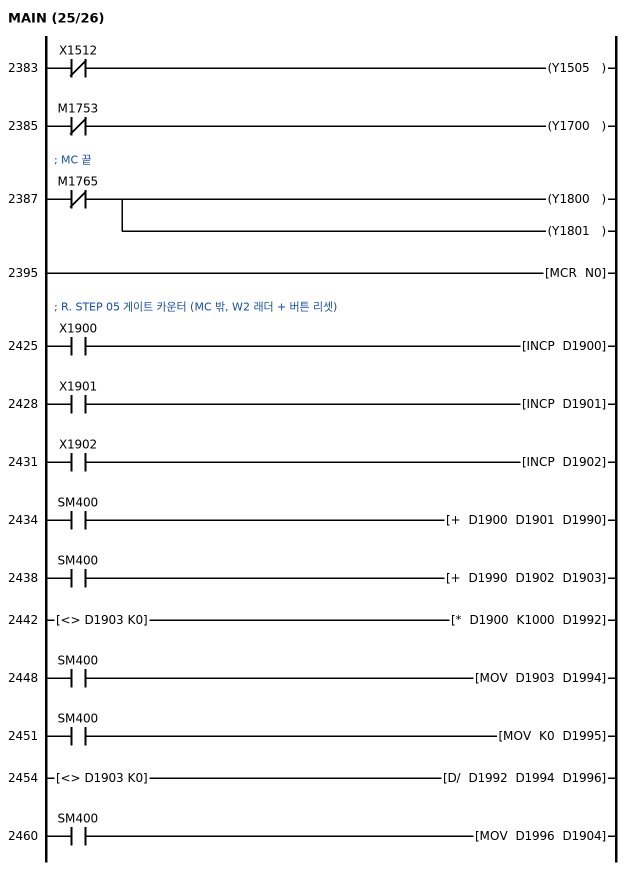
[picture p24: ladder of MAIN, rungs at steps 2383 to 2460]
2383  LDI     X1512
      OUT     Y1505
2385  LDI     M1753
      OUT     Y1700
2387  LDI     M1765
      OUT     Y1800
      OUT     Y1801
; MC 끝
2395  MCR     N0
; R. STEP 05 게이트 카운터 (MC 밖, W2 래더 + 버튼 리셋)
2425  LD      X1900
      INCP    D1900
2428  LD      X1901
      INCP    D1901
2431  LD      X1902
      INCP    D1902
2434  LD      SM400
      +       D1900 D1901 D1990
2438  LD      SM400
      +       D1990 D1902 D1903
2442  LD<>    D1903 K0
      *       D1900 K1000 D1992
2448  LD      SM400
      MOV     D1903 D1994
2451  LD      SM400
      MOV     K0 D1995
2454  LD<>    D1903 K0
      D/      D1992 D1994 D1996
2460  LD      SM400
      MOV     D1996 D1904
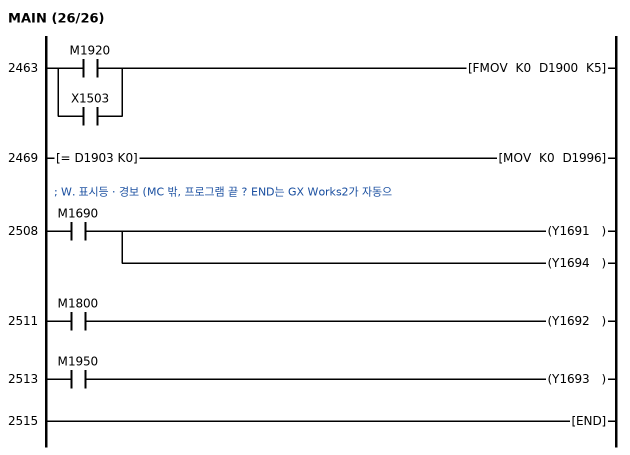
2463  LD      M1920
      OR      X1503
      FMOV    K0 D1900 K5
2469  LD=     D1903 K0
      MOV     K0 D1996
; W. 표시등 · 경보 (MC 밖, 프로그램 끝 ? END는 GX Works2가 자동으
2508  LD      M1690
      OUT     Y1691
      OUT     Y1694
2511  LD      M1800
      OUT     Y1692
2513  LD      M1950
      OUT     Y1693
2515  END
END_PROGRAM
